//{attribute 'qualified_only'}
VAR_GLOBAL	
	fbAnalogSensor			: ARRAY[0..E_ASense_Name.last] OF FB_AnalogSensor;
	
	//arAnalogSensorName		: ARRAY[0..E_ASense_Name.last] OF STRING(12);
	
	//arAnalogSensorRawValue	: ARRAY[0..E_ASense_Name.last] OF INT;

	iAnalogSensor_sel		: INT:=1;
	
	arAnalogSensorNameList	: ARRAY[0..E_ASense_Name.last] OF STRING(12);
	eAnalogSensorNameList	: E_ASense_Name;

	
END_VAR
//{attribute 'qualified_only'}
VAR_GLOBAL PERSISTENT
	//stAnalogSensorSetting	: ARRAY[0..E_Pis_Name.last] OF ST_Piston_Setting_Param;
	stAnalogSensor			: ARRAY[0..E_ASense_Name.last] OF ST_AnalogSensor;
END_VAR

VAR_GLOBAL CONSTANT

END_VAR

(* stored: Version 1.1.0.1, ProductVersion 3.1.4024.12
   GVL g_AnalogSensor: Id {d71deacb-06c5-4b46-a62b-1e15bc291d73} *)
